(* IEC 61131-3 sources: JingjiangArm/moonboxpro_arm_8.4/Application/Application/任务列表/TensionTask/张力控制/收放料/其他, 4 files *)

(* ---- KS_DebugVelCtl.st ---- *)
(*@CES
Name=KS_DebugVelCtl
Type=FunctionBlock
TypeGuid=6f9dac99-8de1-4efc-8465-68ac443b7d08
Guid=5bddb8b6-d642-4e27-baef-5c1f07abfbd7
HasDeclaration=True
HasImplementation=True
*)
{DECLARATION}
FUNCTION KS_DebugVelCtl : BOOL(*调试的速度控制|包含使能标志*)
(*2024.04.12.181136 增加了计算最大加速度的速度输入*)
VAR_INPUT
	i_xDebugEn:BOOL;(*调试使能*)
	i_xRun:BOOL;(*运行标志*)
	i_xStopFast:BOOL;(*快停标志|类似急停时候使能*)
	i_xStopByDec:BOOL;(*减速停止|-TRUE 减速停止|FALSE 直接取消使能停止*)
	i_xManuAcc:BOOL;(*手动加速*)
	i_xManuDec:BOOL;(*手动减速*)
	i_xAutuoAccDec:BOOL;(*自动加减速*)
	i_iVel_Max_mpm:INT;(*最大速度*)
	i_rAxisGirth:REAL;(*轴周长mm*)
	i_rVel_Tar_mpm:REAL;(*目标线速度|m/min*)
	i_pxRunning:POINTER TO BOOL;(*运行中|用来控制使能信号*)
	i_prVel_Cur_mpm:POINTER TO REAL;(*当前线速度|M/MIN*)
	i_prVel_Cur_rpm:POINTER TO REAL;(*当前转速|r/min*)
	i_uiMaxVel_UseCalcAcc:UINT;(*2024.04.12.180908+*)
	i_iCycleTime_Plc: INT;
END_VAR
VAR
	rVel_Cur_mpm:REAL;
	rVel_Cur_rpm:REAL;
	xRunning:BOOL;(*运行中*)
	iAccTime_Nor:INT:=20;(*正常加速时间|S*)
	iDecTime_Nor:INT:=10;(*正常停止时间|S*)
	iDecTime_Fast:INT:=2;(*快停时间|s*)
	iDecTime_Cur: INT;(*当前减速时间*)
	rVel_Tar_mpm: REAL;(*目标速度|输入赋值*)
	rVel_CurTar_mpm: REAL;(*目标速度|=-222为手动加速使能|正常值则为自动加减速*)
	xAutuoAccDec: BOOL;(*自动加减速标志*)
END_VAR
{IMPLEMENTATION}
(*取运行使能*)
IF i_pxRunning<>0 THEN
	xRunning:=i_pxRunning^;
END_IF
(*取线速度和转速*)
IF i_prVel_Cur_mpm<>0 THEN
	rVel_Cur_mpm:=i_prVel_Cur_mpm^;
END_IF
IF i_prVel_Cur_rpm<>0 THEN
	rVel_Cur_rpm:=i_prVel_Cur_rpm^;
END_IF

xAutuoAccDec:=i_xAutuoAccDec;
rVel_Tar_mpm:=i_rVel_Tar_mpm;

iDecTime_Cur:=iDecTime_Nor;
IF i_xStopFast THEN
	iDecTime_Cur:=iDecTime_Fast;
END_IF

(*执行部分*)
IF i_xDebugEn THEN(*调试使能|*)
	(*使能标志处理*)
	IF i_xRun THEN(*运行有效*)
		IF NOT xRunning THEN(*非运行中*)
			xRunning:=TRUE;(*输出运行中标志|控制电机使能*)
		END_IF
	END_IF
END_IF

(*停止是标志处理|*)
IF NOT i_xDebugEn OR
	NOT i_xRun THEN
	IF NOT i_xStopByDec THEN
		xRunning:=FALSE;
		rVel_Cur_mpm:=0.0;(*速度写0*)
	ELSE(*停止到0*)
		IF rVel_Cur_mpm>=0.0001 THEN
			xAutuoAccDec:=TRUE;
			rVel_Tar_mpm:=0;
		END_IF
	END_IF

	IF rVel_Cur_mpm<=0.0001 THEN(*用线速度作为条件*)
		xRunning:=FALSE;
		rVel_Cur_mpm:=0.0;(*速度写0*)
	END_IF
END_IF
(*自动加减速控制|*)
IF xAutuoAccDec THEN
	rVel_CurTar_mpm:=rVel_Tar_mpm;
ELSE(**非自动加减速*)
	rVel_Tar_mpm:=-222;
END_IF

KS_VelPrf(
	xRunning,
	i_xManuAcc,
	i_xManuDec,
	i_iCycleTime_Plc,
	iAccTime_Nor,
	iDecTime_Cur,
	i_iVel_Max_mpm,
	rVel_Tar_mpm,
	ADR(rVel_Cur_mpm),
	i_uiMaxVel_UseCalcAcc);(*2024.04.12.181005+*)

(*将线速度转换为转速*)
IF i_rAxisGirth<>0 THEN
	rVel_Cur_rpm:=rVel_Cur_mpm*1000/i_rAxisGirth;
ELSE
	rVel_Cur_rpm:=0;
END_IF

(*取运行使能*)
IF i_pxRunning<>0 THEN
	i_pxRunning^:=xRunning;
END_IF
(*输出线速度和转速*)
IF i_prVel_Cur_mpm<>0 THEN
	i_prVel_Cur_mpm^:=rVel_Cur_mpm;
END_IF
IF i_prVel_Cur_rpm<>0 THEN
	i_prVel_Cur_rpm^:=rVel_Cur_rpm;
END_IF

(* ---- KS_GetMax_MinVlaue.st ---- *)
(*@CES
Name=KS_GetMax_MinVlaue
Type=FunctionBlock
TypeGuid=6f9dac99-8de1-4efc-8465-68ac443b7d08
Guid=8f6e33c8-95eb-4af2-849c-6572b367cef7
HasDeclaration=True
HasImplementation=True
*)
{DECLARATION}
FUNCTION KS_GetMax_MinVlaue : INT(*获取最大或者最小值*)
VAR_INPUT
	i_plrMaxValue:POINTER TO LREAL;(*大值*)
	i_plrMinValue:POINTER TO LREAL;(*小值*)
	i_lrValue:LREAL;(*值*)
END_VAR
VAR
END_VAR
{IMPLEMENTATION}
KS_GetMax_MinVlaue:=0;
IF i_plrMaxValue<>0 AND i_plrMinValue<>0 THEN
	IF i_lrValue>i_plrMaxValue^ THEN
		i_plrMaxValue^:=i_lrValue;
	ELSIF i_lrValue<i_plrMinValue^ THEN
		i_plrMinValue^:=i_lrValue;
	ELSE;
	END_IF
ELSE
	KS_GetMax_MinVlaue:=-1;
END_IF

(* ---- KS_VelPrf.st ---- *)
(*@CES
Name=KS_VelPrf
Type=FunctionBlock
TypeGuid=6f9dac99-8de1-4efc-8465-68ac443b7d08
Guid=b931f0d4-2560-4387-b073-ed705f607109
HasDeclaration=True
HasImplementation=True
*)
{DECLARATION}
FUNCTION KS_VelPrf : BOOL
(*2024.04.12.181136 增加了计算最大加速度的速度输入*)
VAR_INPUT
	i_xEn:BOOL;(*规划使能*)
	i_xAcc:BOOL;(*加速*)
	i_xDec:BOOL;(*减速*)
	i_iTime_PlcCycle:INT:=20;(*plc执行时间*)
	i_iAccTime:INT;(*加速时间S|0加速到最大速度的时间|写0则直接赋值*)
	i_iDecTime:INT;(*减速时间S|由最大速度减速到0的时间|写0则直接赋值*)
	i_iVel_Max:INT;(*最大速度|用来计算加速度*)
	i_rVel_Tar:REAL;(*目标速度|如果目标速度等于特殊值 例如-222，我们根据按钮加减速。否则根据目标速度加减速*)
	i_prVel_Cur:POINTER TO REAL;(*当前速度*)
	i_uiMaxVel_UseCalcAcc:UINT;(*2024.04.12.180908+*)
END_VAR
VAR
	lrAcceleration: LREAL;(*加速度|m/min/ms*)
	lrDeceleration: LREAL;(*减加速度|m/min/ms*)
	xAcc: BOOL;
	xDec: BOOL;
	lrVel_Tar: LREAL;(*目标速度*)
END_VAR
{IMPLEMENTATION}
IF i_xEn THEN(*规划使能*)
	IF  i_prVel_Cur<>0 THEN
		(*计算加减速度*)
		IF i_iAccTime>0 THEN
			lrAcceleration:=UINT_TO_LREAL(i_uiMaxVel_UseCalcAcc)/i_iAccTime/1000;(*加速度*)
		END_IF
		IF i_iDecTime>0 THEN
			lrDeceleration:=-UINT_TO_LREAL(i_uiMaxVel_UseCalcAcc)/i_iDecTime/1000;(*减加速度*)
		END_IF

		lrVel_Tar:=i_rVel_Tar;
		(*判断加减速状态*)
		IF i_rVel_Tar<>-222 THEN(*根据目标速度确定加减速*)
			IF i_prVel_Cur^>i_rVel_Tar THEN
				xDec:=TRUE;
			ELSIF i_prVel_Cur^<i_rVel_Tar THEN
				xAcc:=TRUE;
			END_IF
		ELSE(*根据按钮确定加减速度*)
			xAcc:=i_xAcc;(*按钮同时按下 则是加速*)
			xDec:=NOT xAcc AND i_xDec;

			IF xAcc THEN(*加速我们加到最大速度*)
				lrVel_Tar:=i_iVel_Max;
			ELSIF xDec THEN(*减速我们减到0*)
				lrVel_Tar:=0;
			END_IF
		END_IF

		IF xAcc THEN(*加速*)
			IF lrAcceleration<>0 THEN
				i_prVel_Cur^:=i_prVel_Cur^+LREAL_TO_REAL(lrAcceleration*i_iTime_PlcCycle);
				IF i_prVel_Cur^>lrVel_Tar THEN
					i_prVel_Cur^:=LREAL_TO_REAL(lrVel_Tar);
				END_IF
			ELSE
				i_prVel_Cur^:=LREAL_TO_REAL(lrVel_Tar);
			END_IF
		ELSIF xDec THEN(*减速*)
			IF lrDeceleration<>0 THEN
				i_prVel_Cur^:=i_prVel_Cur^+LREAL_TO_REAL(lrDeceleration*i_iTime_PlcCycle);
				IF i_prVel_Cur^<lrVel_Tar THEN
					i_prVel_Cur^:=LREAL_TO_REAL(lrVel_Tar);
				END_IF
			ELSE
				i_prVel_Cur^:=LREAL_TO_REAL(lrVel_Tar);
			END_IF
		END_IF
	END_IF
ELSE(*规划取消*)
	i_prVel_Cur^:=0;
END_IF

(* ---- KS_FB_AxisDebug.st ---- *)
(*@CES
Name=KS_FB_AxisDebug
Type=FunctionBlock
TypeGuid=6f9dac99-8de1-4efc-8465-68ac443b7d08
Guid=225e022e-2ac6-4e18-87bd-0bf6abe85a88
HasDeclaration=True
HasImplementation=True
*)
{DECLARATION}
FUNCTION_BLOCK KS_FB_AxisDebug
VAR_INPUT
	i_xEn:BOOL;
	i_xEstopBtn:BOOL;(*急停*)
	i_xFlag_Estop: BOOL;
	i_xFlag_Tension: BOOL;
	i_xFlag_Print: BOOL;
	i_xCurAxisA: BOOL;
	i_rVel_Max: REAL;
	i_xFuncBtn:BOOL;(*放料功能按钮|单击-根据当前轴选择控制加速哪一个轴|延迟1s后加速-考虑使用伺服初始化耗时-接料准备时候不能按钮不能使用了
									  双击(500MS内按下2次)-控制停止ab轴|
									  常按3s则根据当前轴选择控制停止哪一个轴*)
	(*2021.10.14.102041*)
	i_xPreCutBtn:BOOL;(*接料准备*)
	i_xCutCancelBtn:BOOL;(*接料解除-退出接料准备状态并减速*)
	i_xCutBtn:BOOL;(*接料|单击是接料|双击则自动加速到目标速度或者停止到当前速度*)
	i_xStsPreCut:BOOL;(*接料准备状态*)
	i_iDebugVelmpm_AxisA:INT;(*A轴调试速度|m/min*)
	i_iDebugGirthmm_AxisA:INT;(*调试的A轴周长*)
	i_iDebugVelmpm_AxisB:INT;(*B轴调试速度|m/min*)
	i_iDebugGirthmm_AxisB:INT;(*调试的B轴周长*)
	i_iCycleTime_Plc: INT;
END_VAR
VAR_OUTPUT
	o_xEn:BOOL;
	o_xLampFlick_Debug:BOOL;(*指示调试预驱同步有效标志-加减速250MS闪烁|处于调试状态*)
	(*接料准备动作逻辑兼容|2021.10.14.101833*)
	o_xPreCut_Debug:BOOL;(*接料准备调试按钮输出*)
	o_xCutCancel_Debug:BOOL;(*接料取消调试按钮输出|可能不需要*)
	o_xCut_Debug:BOOL;(*接料调试按钮输出*)
	o_xLamp_PreDrive_Debug:BOOL;(*调试预驱同步输出*)
END_VAR
VAR
	xStopFast:BOOL;(*快停|用于处理急停*)
	xFlag_NeedStop: BOOL;(*停止标志*)
	xAxisDebugEn: BOOL;(*放料轴调试使能|.0*)
	xAxisADebugRun: BOOL;(*放料A轴调试运行|.1*)
	xAxisADebugAutoAccDec: BOOL;(*放料A轴调试自动加减速|.2*)
	xAxisADebugRunning: BOOL;(*放料A轴调试运行中|作为输出|.3*)
	xAxisBDebugRun: BOOL;(*放料B轴调试运行|.4*)
	xAxisBDebugAutoAccDec: BOOL;(*放料B轴调试自动加减速|.5*)
	xAxisBDebugRunning: BOOL;(*放料B轴调试运行中|作为输出|.6*)
	xLastFuncBtn:BOOL;(*功能键按下上个周期值*)
	tTimeFuncBtnDn: TIME;(*放料功能键按下时间|按下沿的时间*)
	iClickNum: BYTE;(*点击次数*)
	tTimeRetain:TIME:=T#3S;(*放料功能键按下持续时间时间|按下超过这个时间就只停止a\b轴*)
	tTimeDoubleClick:TIME:=T#500MS;(*放料功能键按下单双击时间|*)
	tDelayTimeAutoAccByBtn:TIME:=T#1S;(*放料通过放料面板自动加速延迟时间*)
	xAllAxisStop: BOOL;(*ab轴都停止标志*)
	fbAxisAStopTrig:R_TRIG;(*放料A轴停止沿*)
	fbAxisBStopTrig:R_TRIG;(*放料B轴停止沿*)
	xAxisAStop: BOOL;(*a轴停止标志*)
	xAxisBStop: BOOL;(*b轴停止标志*)
	xAxisAAutoAcc: BOOL;(*A轴自动加速标志*)
	fbTon_AxisAAutoAcc: TON;(*A轴自动加速延时器*)
	fbRTrig_AxisAAutoAcc: R_TRIG;(*A轴自动加速沿*)
	xAxisBAutoAcc: BOOL;(*B轴自动加速标志*)
	fbTon_AxisBAutoAcc: TON;(*B轴自动加速延时器*)
	fbRTrig_AxisBAutoAcc: R_TRIG;(*B轴自动加速沿*)
	xAxisAccOrDecing:BOOL;(*放料变速状态中*)
	fbTon_AxisAccOrDecingFlick: TON;(*轴加减速中闪烁计时器*)
	xLampFlick_Debug:BOOL;(*闪烁指示灯*)

	afbTrigBtn:ARRAY [1..3] OF R_TRIG;
	xReqPreCut: BOOL;(*接料准备沿*)
	xReqCutCancel: BOOL;(*接料取消沿*)
	xReqCut: BOOL;(*接料沿*)
	iCutBtnClickNum: INT;
	tTimeCutBtnDn: TIME;
	xLastStsPreCut:BOOL;
	xAxisDebuging: BOOL;(*调试中标志*)
	rAxisAVelTar: REAL;(*A轴目标速度*)
	rAxisBVelTar: REAL;(*B轴目标速度*)
	arLastCurVel: ARRAY [1..4] OF REAL;(*收放料4个轴的速度备份|判断在变速状态*)
END_VAR
VAR_IN_OUT
	io_xAxisDebugEn: BOOL;
	io_xAxisADebugRun: BOOL;
	io_xAxisBDebugRun: BOOL;
	io_xAxisADebugRunning: BOOL;
	io_xAxisBDebugRunning: BOOL;
	io_xAxisADebugAutoAccDec: BOOL;
	io_xAxisBDebugAutoAccDec: BOOL;

	io_rDebugCurVelmpmAxisA: REAL;
	io_rDebugCurVelmpmAxisB: REAL;
	io_rDebugCurVelrpmAxisA: REAL;
	io_rDebugCurVelrpmAxisB: REAL;
END_VAR
{IMPLEMENTATION}
xAxisDebugEn:=io_xAxisDebugEn;
(*放料A轴测试|*)
IF io_rDebugCurVelmpmAxisA=0 THEN
	xAxisADebugRun:=io_xAxisADebugRun;
ELSE
	IF NOT io_xAxisADebugRun THEN
		xAxisADebugRun:=io_xAxisADebugRun;
	END_IF
END_IF
xAxisADebugAutoAccDec:= io_xAxisADebugAutoAccDec;
(*放料b轴测试*)
IF io_rDebugCurVelmpmAxisB=0 THEN
	xAxisBDebugRun:=io_xAxisBDebugRun;
ELSE
	IF NOT io_xAxisBDebugRun THEN
		xAxisBDebugRun:=io_xAxisBDebugRun;
	END_IF
END_IF
xAxisBDebugAutoAccDec:=io_xAxisBDebugAutoAccDec;
(*数值合法性处理*)
IF i_iDebugGirthmm_AxisA=0 THEN i_iDebugGirthmm_AxisA:=300;END_IF
IF i_iDebugVelmpm_AxisA=0 THEN i_iDebugVelmpm_AxisA:=300;END_IF
IF i_iDebugGirthmm_AxisB=0 THEN i_iDebugGirthmm_AxisB:=300;END_IF
IF i_iDebugVelmpm_AxisB=0 THEN i_iDebugVelmpm_AxisB:=300;END_IF

IF i_xEstopBtn OR i_xFlag_Estop  THEN
	xStopFast:=TRUE;(*急停时候使用快速停止*)
	xFlag_NeedStop:=TRUE;
ELSE
	IF xFlag_NeedStop THEN
		IF NOT (xAxisADebugRunning OR
			xAxisBDebugRunning) THEN(*所有轴都停止使能了|复位标志*)
			xStopFast:=FALSE;
			xFlag_NeedStop:=FALSE;
		END_IF
	END_IF
END_IF

(*针对收放料的处理*)
IF  xFlag_NeedStop OR (*急停的时候需要停止运动*)
	i_xFlag_Tension OR(*使用收放料的时候就停止调试*)
(*		i_pstStGrpParam^.xFlag_Ink or(*空转 我们认为是开机|就停止调试*)*)
	i_xFlag_Print THEN(*印刷时候|就停止调试|2022.4.10.154641*)
	(*放料A轴清除*)
	xAxisADebugRun:=FALSE;
	xAxisAAutoAcc:=FALSE;
	xAxisADebugAutoAccDec:=FALSE;
	(*放料B轴清除*)
	xAxisBDebugRun:=FALSE;
	xAxisBAutoAcc:=FALSE;
	xAxisBDebugAutoAccDec:=FALSE;

	IF NOT xFlag_NeedStop THEN(*不是急停停止的时候我们退出调试模式|*)
		xAxisDebugEn:=FALSE;
		xAxisDebugEn:=FALSE;
	END_IF
END_IF

(****************************************************************************************************)
xAllAxisStop:=FALSE;
xAxisAStop:=FALSE;
xAxisBStop:=FALSE;
(*接料准备动作逻辑兼容|2021.10.14.101833*)
o_xPreCut_Debug:=FALSE;(*接料准备调试按钮输出*)
o_xCutCancel_Debug:=FALSE;(*接料取消调试按钮输出|可能不需要*)
o_xCut_Debug:=FALSE;(*接料调试按钮输出*)
o_xLamp_PreDrive_Debug:=FALSE;
(*放料轴停止\加速|*)
afbTrigBtn[1](CLK:=i_xPreCutBtn,Q=>xReqPreCut);
afbTrigBtn[2](CLK:=i_xCutCancelBtn,Q=>xReqCutCancel);
afbTrigBtn[3](CLK:=i_xCutBtn,Q=>xReqCut);
IF xAxisDebugEn THEN
	xAxisDebuging:=TRUE;
	(*2021.10.14.110723 兼容的接料准备逻辑------------------------------------------*)
	IF xReqPreCut AND NOT i_xStsPreCut THEN(*接料准备*)
		o_xPreCut_Debug:=TRUE;
	END_IF
	IF i_xStsPreCut THEN(*进入接料准备时候常输出运动使能标志*)
		IF io_rDebugCurVelmpmAxisA=0 THEN
			xAxisADebugRun:=TRUE;(*使能启动*)
		END_IF
		IF io_rDebugCurVelmpmAxisB=0 THEN
			xAxisBDebugRun:=TRUE;(*使能启动*)
		END_IF

		IF i_xCurAxisA THEN(*A轴|B轴常输出加速状态|下面当前速度会根据A轴速度改变*)
			xAxisBAutoAcc:=xAxisBDebugRun;
		ELSE
			xAxisAAutoAcc:=xAxisADebugRun;
		END_IF

		IF io_rDebugCurVelmpmAxisA = io_rDebugCurVelmpmAxisB AND
			io_rDebugCurVelmpmAxisA<>0 THEN(*调试速度相等|并且不等于0 认为同步了*)
			o_xLamp_PreDrive_Debug:=TRUE;
		END_IF
		(*接料准备情况下不考虑功能按键|2021.10.14.102751
		控制由接料准备和接料解除接管*)
		i_xFuncBtn:=FALSE;
		IF xReqCut THEN
			iCutBtnClickNum:=iCutBtnClickNum+1;
			IF iCutBtnClickNum=1 THEN
				tTimeCutBtnDn:=TIME();
			END_IF
		END_IF
		IF iCutBtnClickNum>=2 THEN(*按下2次|加速或者停止*)
			iCutBtnClickNum:=0;
			IF i_xCurAxisA THEN(*A轴*)
				xAxisAAutoAcc:=NOT xAxisAAutoAcc;
			ELSE
				xAxisBAutoAcc:=NOT xAxisBAutoAcc;
			END_IF
		ELSE
			(*超过500MS未再次按下|我们认为是单击事件|根据当前轴切换自动加速*)
			IF iCutBtnClickNum>0 THEN(*已经按下了|启动计时，如果500MS内未再次按下，则清除计数*)
				IF TIME()-tTimeCutBtnDn>=tTimeDoubleClick THEN
					o_xCut_Debug:=o_xLamp_PreDrive_Debug AND NOT xAxisAccOrDecing;(*预驱同步了不在加减速才能输出裁切*)
					iCutBtnClickNum:=0;
				END_IF
			END_IF
		END_IF

		IF xReqCutCancel THEN(*接料解除|并停止速度*)
			o_xCutCancel_Debug:=TRUE;
			xAllAxisStop:=TRUE;
		END_IF
	ELSE
		IF xLastStsPreCut THEN(*退出接料状态了|全体停止*)
			xAllAxisStop:=TRUE;
		END_IF
		iCutBtnClickNum:=0;
	END_IF
	(*2021.10.14.110723 兼容的接料准备逻辑------------------------------------------*)

	IF i_xFuncBtn AND NOT xLastFuncBtn THEN(*停止|*)
		iClickNum:=iClickNum+1;
		IF iClickNum=1 THEN
			tTimeFuncBtnDn:=TIME();
		END_IF
	END_IF

	IF iClickNum>=2 THEN(*按下2次|ab轴停止*)
		iClickNum:=0;
		xAllAxisStop:=TRUE;
	ELSE
		(*超过500MS未再次按下|我们认为是单击事件|根据当前轴切换自动加速*)
		IF iClickNum>0 THEN(*已经按下了|启动计时，如果500MS内未再次按下，则清除计数*)
			IF TIME()-tTimeFuncBtnDn>=tTimeDoubleClick THEN
				IF NOT i_xFuncBtn THEN(*超过tTimeDoubleClick_Uw按钮也抬起来了|*)
					IF i_xCurAxisA THEN(*A轴*)
						IF io_rDebugCurVelmpmAxisA=0 THEN
							xAxisADebugRun:=TRUE;(*使能启动*)
						END_IF
						IF xAxisADebugRun THEN
							xAxisAAutoAcc:=NOT xAxisAAutoAcc;
						END_IF
					ELSE(**B轴*)
						IF io_rDebugCurVelmpmAxisB=0 THEN
							xAxisBDebugRun:=TRUE;(*使能启动*)
						END_IF
						IF xAxisBDebugRun THEN
							xAxisBAutoAcc:=NOT xAxisBAutoAcc;
						END_IF
					END_IF
				END_IF
				iClickNum:=0;
			END_IF
		END_IF
	END_IF

	IF i_xFuncBtn THEN(*常按下|根据当前轴 分轴停止*)
		IF TIME()-tTimeFuncBtnDn>=tTimeRetain THEN
			IF i_xCurAxisA THEN(*A轴*)
				xAxisAStop:=TRUE;
			ELSE(**B轴*)
				xAxisBStop:=TRUE;
			END_IF
		END_IF
	END_IF

	fbAxisAStopTrig(CLK:=xAxisAStop);
	fbAxisBStopTrig(CLK:=xAxisBStop);
	IF fbAxisAStopTrig.Q OR
		fbAxisBStopTrig.Q OR
		xAllAxisStop  THEN
		(*放料A轴清除*)
		IF xAxisAStop OR xAllAxisStop THEN
			xAxisADebugRun:=FALSE;
			xAxisAAutoAcc:=FALSE;
			xAxisADebugAutoAccDec:=FALSE;
		END_IF
		(*放料B轴清除*)
		IF xAxisBStop OR xAllAxisStop THEN
			xAxisBDebugRun:=FALSE;
			xAxisBAutoAcc:=FALSE;
			xAxisBDebugAutoAccDec:=FALSE;
		END_IF
	END_IF

	(*延时自动加速*)
	IF NOT xAxisAAutoAcc AND fbTon_AxisAAutoAcc.IN THEN(*取消自动加速|复位标志*)
		xAxisADebugAutoAccDec:=FALSE;
	END_IF
	fbTon_AxisAAutoAcc(IN:=xAxisAAutoAcc,PT:=T#1S);
	fbRTrig_AxisAAutoAcc(CLK:=fbTon_AxisAAutoAcc.Q);
	IF fbRTrig_AxisAAutoAcc.Q THEN(*延时1s加速|考虑到收放料使用伺服情况下的初始化动作时间*)
		xAxisADebugAutoAccDec:=TRUE;
	END_IF
	(*在关闭运动使能的时候清除自动加减速标志*)
	(*没有使能的时候关闭自动减速*)
	IF NOT xAxisADebugRun THEN
		xAxisADebugAutoAccDec:=FALSE;
	END_IF
	(*延时自动加速*)
	IF NOT xAxisBAutoAcc AND fbTon_AxisBAutoAcc.IN THEN(*取消自动加速|复位标志*)
		xAxisBDebugAutoAccDec:=FALSE;
	END_IF
	fbTon_AxisBAutoAcc(IN:=xAxisBAutoAcc,PT:=tDelayTimeAutoAccByBtn);
	fbRTrig_AxisBAutoAcc(CLK:=fbTon_AxisBAutoAcc.Q);
	IF fbRTrig_AxisBAutoAcc.Q THEN(*延时1s加速|考虑到收放料使用伺服情况下的初始化动作时间*)
		xAxisBDebugAutoAccDec:=TRUE;
	END_IF
	(*在关闭运动使能的时候清除自动加减速标志*)
	(*没有使能的时候关闭自动减速*)
	IF NOT xAxisBDebugRun THEN
		xAxisBDebugAutoAccDec:=FALSE;
	END_IF
ELSE(*非调试模式*)
	IF xAxisDebuging THEN(*调试中|如果有接料准备则退出*)
		xAxisDebuging:=FALSE;
		IF i_xStsPreCut THEN
			o_xCutCancel_Debug:=TRUE;
		END_IF
	END_IF
	iClickNum:=0;
	fbAxisAStopTrig(CLK:=FALSE);
	fbAxisBStopTrig(CLK:=FALSE);
	fbTon_AxisAAutoAcc(IN:=FALSE);
	fbRTrig_AxisAAutoAcc(CLK:=FALSE);
	fbTon_AxisBAutoAcc(IN:=FALSE);
	fbRTrig_AxisBAutoAcc(CLK:=FALSE);
	xAxisADebugRun:=FALSE;
	xAxisADebugAutoAccDec:=FALSE;
	xAxisBDebugRun:=FALSE;
	xAxisBDebugAutoAccDec:=FALSE;
	xAxisAAutoAcc:=FALSE;
	xAxisBAutoAcc:=FALSE;
END_IF
xLastFuncBtn:=i_xFuncBtn;
xLastStsPreCut:=i_xStsPreCut;

(*放A速度控制*)
rAxisAVelTar:=i_iDebugVelmpm_AxisA;
IF i_xStsPreCut THEN(*接料准备状态下|目标速度为当前轴的速度*)
	IF i_xCurAxisA THEN(*当前轴是A轴*);
	ELSE(*当前轴B轴|A轴的目标速度=B轴当前速度*)
		rAxisAVelTar:=io_rDebugCurVelmpmAxisB;
	END_IF
END_IF

KS_DebugVelCtl(
	xAxisDebugEn,
	xAxisADebugRun,
	xStopFast,
	TRUE,
	FALSE,
	FALSE,
	xAxisADebugAutoAccDec,
	LREAL_TO_INT(i_rVel_Max),
	i_iDebugGirthmm_AxisA,
	rAxisAVelTar,
	ADR(xAxisADebugRunning),
	ADR(io_rDebugCurVelmpmAxisA),
	ADR(io_rDebugCurVelrpmAxisA),
	LREAL_TO_UINT(i_rVel_Max),
	i_iCycleTime_Plc);(*2024.04.12.181058+*)

(*放B速度控制*)
rAxisBVelTar:=i_iDebugVelmpm_AxisB;
IF i_xStsPreCut THEN(*接料准备状态下|目标速度为当前轴的速度*)
	IF i_xCurAxisA THEN(*当前轴是A轴|B轴的目标速度=A轴当前速度*);
		rAxisBVelTar:=io_rDebugCurVelmpmAxisA;
	ELSE(*当前轴B轴|A轴的目标速度=B轴当前速度*);
	END_IF
END_IF

KS_DebugVelCtl(
	xAxisDebugEn,
	xAxisBDebugRun,
	xStopFast,
	TRUE,
	FALSE,
	FALSE,
	xAxisBDebugAutoAccDec,
	LREAL_TO_INT(i_rVel_Max),
	i_iDebugGirthmm_AxisB,
	rAxisBVelTar,
	ADR(xAxisBDebugRunning),
	ADR(io_rDebugCurVelmpmAxisB),
	ADR(io_rDebugCurVelrpmAxisB),
	LREAL_TO_UINT(i_rVel_Max),
	i_iCycleTime_Plc);(*2024.04.12.181058+*)

(****************************************************************************************************)

xAxisAccOrDecing:=FALSE;
IF arLastCurVel[1]<>io_rDebugCurVelmpmAxisA OR
	arLastCurVel[2]<>io_rDebugCurVelmpmAxisB THEN
	xAxisAccOrDecing:=TRUE;
END_IF

arLastCurVel[1]:=io_rDebugCurVelmpmAxisA;
arLastCurVel[2]:=io_rDebugCurVelmpmAxisB;

(*调试模式指示灯闪烁指示*)
fbTon_AxisAccOrDecingFlick(IN:=xAxisAccOrDecing,PT:=T#250MS);
IF fbTon_AxisAccOrDecingFlick.Q THEN(*加减速中使用500ms闪烁指示|*)
	xLampFlick_Debug:=NOT xLampFlick_Debug;
	fbTon_AxisAccOrDecingFlick(IN:=FALSE);
ELSIF NOT xAxisAccOrDecing THEN(*停止加减速|输出同步指示*)
	xLampFlick_Debug:=o_xLamp_PreDrive_Debug;
END_IF
o_xLampFlick_Debug:=xAxisDebugEn AND xLampFlick_Debug;
(*放料调试模式*)
(*i_pstStGrpParam^.wAxisDebug_UwRw.0*)
io_xAxisDebugEn :=xAxisDebugEn;
(*放料A*)
(*i_pstStGrpParam^.wAxisDebug_UwRw.1*)
io_xAxisADebugRun:=xAxisADebugRun;
(*i_pstStGrpParam^.wAxisDebug_UwRw.2*)
io_xAxisADebugAutoAccDec:=xAxisADebugAutoAccDec;
(*i_pstStGrpParam^.wAxisDebug_UwRw.3*)
io_xAxisADebugRunning:=xAxisADebugRunning;
(*放料B*)
(*i_pstStGrpParam^.wAxisDebug_UwRw.4*)
io_xAxisBDebugRun:=xAxisBDebugRun;
(*i_pstStGrpParam^.wAxisDebug_UwRw.5*)
io_xAxisBDebugAutoAccDec:=xAxisBDebugAutoAccDec;
(*i_pstStGrpParam^.wAxisDebug_UwRw.6*)
io_xAxisBDebugRunning:=xAxisBDebugRunning;

o_xEn:=i_xEn;
